PROGRAM MAIN
VAR
	fbIgorCtrl:			FB_IgorCtrl;
END_VAR

fbIgorCtrl();

END_PROGRAM

(* stored: Version 1.1.0.1, ProductVersion 3.1.4024.9
   POU MAIN: Id {8fb21f47-0787-4c92-8c3b-9716b5a9abe0}, SpecialFunc None *)
